{attribute 'qualified_only'}
VAR_GLOBAL
    // Operator / HMI / sequence commands (internal PLC tags)
    bEStop1_ResetCmd     : BOOL;         // Momentary reset request from HMI/button
    bSafety_ErrAckCmd    : BOOL;         // Momentary error acknowledge request

    // Rising-edge outputs mapped to TwinSAFE standard aliases (PLC -> TwinSAFE)
    bEStop1_RestartOut   AT %Q* : BOOL;  // Linked to EStop1_Restart.sds
    bSafety_ErrAckOut    AT %Q* : BOOL;  // Linked to ErrorAcknowledgement.sds
    bSafety_GroupRunOut  AT %Q* : BOOL;  // Linked to Run.sds (TwinSAFE group run enable)

    // Safety status & diagnostics (TwinSAFE / I/O -> PLC)
    bEStop1_SafeHealthy  AT %I* : BOOL;  // TRUE when E-Stop safe output is healthy
    bEStop1_Tripped      : BOOL;         // Derived: TRUE when E-Stop is open/tripped
    bSafety_ComFault     AT %I* : BOOL;  // Safety communication / group fault status
END_VAR

(* stored: Version 1.1.0.1
   GVL GVL_Safety: Id {cf88dd38-b736-4d97-b024-1f3ef90e1e6e} *)
